Yaskawa INFORM job: 20211127CHUFENGKOUCOR.JBI

/JOB
//NAME 20211127CHUFENGKOUCOR
//POS
///NPOS 5,0,5,1,0,1
///TOOL 1
///POSTYPE PULSE
///PULSE
C00000=-5456,29378,14097,-3416,-76919,3294
C00001=-6880,32387,-10693,-3890,-57663,4370
C00002=-5335,32532,-16573,-4114,-53450,4057
C00003=-5253,34423,-13635,-4085,-54045,4006
C00004=-5387,38273,25473,-3407,-78050,3239
///TOOL 0
EC00000=-4,321083
EC00001=-4,321083
EC00002=-4,221835
EC00003=-4,93195
EC00004=-4,93198
///TOOL 1
///POSTYPE ROBOT
///RECTAN
///RCONF 0,0,0,0,0,0,0,0,0,0,0,0,0,0,0,0,0,0,0,0,0,0,0,0
P00001=629.883,8.042,-21.694,-154.9112,52.6025,29.7528
///POSTYPE PULSE
///PULSE
EX00001=2,-321071
//INST
///DATE 2021/11/27 15:41
///ATTR SC,RW
///GROUP1 RB1
///GROUP2 ST1
NOP
MOVJ C00000 VJ=10.00  +MOVJ EC00000 VJ=10.00
MOVJ C00001 VJ=10.00  +MOVJ EC00001 VJ=0.78
CALL JOB:STARTDETPRG
WAIT B005=1
MOVL P001 V=10.0  +MOVJ EX001
CALL JOB:ENDDETPRG
CALL JOB:STARTCOR
ARCON AC=160 AV=30.0
SMOVC P001 V=5.0  +MOVJ EX001
SMOVC C00002 V=4.5  +MOVJ EC00002
SMOVC C00003 V=4.5  +MOVJ EC00003
CALL JOB:ENDDETPRG
ARCOF
MOVL C00004 V=20.0  +MOVJ EC00004 VJ=10.00
END
